Fanuc KAREL source: kt00225.KL

-- PROVISIONAL review KL for V940-1; original PC SHA256 ac3c03bb982a2ed19b04aea069ecc35dc1cdea4b9b8599c1d20720946dc370e8
-- Incomplete behavior may be omitted. Consult companion uncertainty JSON. Do not deploy.
PROGRAM KT00225
%NOLOCKGROUP
VAR
  B1 : BOOLEAN
  B2 : BOOLEAN
  OUT : BOOLEAN
BEGIN
  B1 = TRUE
  B2 = FALSE
  B1 = TRUE
  B2 = FALSE
  OUT = (B1 OR B2)
END KT00225
